// TIA Portal V19 export
// export: Created 2026-10-15T10:10:37.1458644Z, ExportSetting WithDefaults, DisplayName Totally Integrated Automation Portal, DisplayVersion V19, DisplayName TIA Portal Openness, DisplayVersion V19, DisplayName TIA Portal Version Control Interface, DisplayVersion V19, DisplayName STEP 7 Professional, DisplayVersion V19, DisplayName STEP 7 Safety, DisplayVersion V19, DisplayName WinCC Basic/Comfort/Advanced, DisplayVersion V19, DisplayName WinCC Unified, DisplayVersion V19
FUNCTION "ROLL_ReadInputs" : Void   // FC36, SCL
{ S7_Optimized_Access := 'TRUE' }
VERSION : 0.1
// stored: AutoNumber true, IsIECCheckEnabled false, SetENOAutomatically false, UDAEnableTagReadback false
   VAR_TEMP
      "b" : Int;
      bit : Int;
   END_VAR
BEGIN

   // Confirmed four-station profile: absent optional inputs are zero.
   FOR #b := 119 TO 125 DO
       FOR #bit := 0 TO 7 DO
           "ROLL_IO".Input[#b, #bit] := FALSE;
       END_FOR;
   END_FOR;
   IF "ROLL_IO".PhysicalIoConfigured AND NOT "ROLL_IO".Simulation THEN
       "ROLL_IO".Input[0, 0] := "Tag__639276557951123186";
       "ROLL_IO".Input[0, 1] := "Tag__639276557952818668";
       "ROLL_IO".Input[0, 2] := "Tag__639276557952918398";
       "ROLL_IO".Input[0, 3] := "Tag__639276557952998183";
       "ROLL_IO".Input[0, 4] := "Tag__639276557953077986";
       "ROLL_IO".Input[0, 5] := "Tag__639276557953157762";
       "ROLL_IO".Input[0, 6] := "Tag__639276557953227573";
       "ROLL_IO".Input[0, 7] := "Tag__639276557953307358";
       "ROLL_IO".Input[1, 0] := "Tag__639276557953367206";
       "ROLL_IO".Input[1, 1] := "Tag__639276557953447409";
       "ROLL_IO".Input[1, 2] := "Tag__639276557953526828";
       "ROLL_IO".Input[1, 3] := "Tag__639276557953606562";
       "ROLL_IO".Input[1, 4] := "Tag__639276557953686353";
       "ROLL_IO".Input[1, 5] := "Tag__639276557953766129";
       "ROLL_IO".Input[1, 6] := "Tag__639276557953835956";
       "ROLL_IO".Input[1, 7] := "Tag__639276557953915729";
       "ROLL_IO".Input[2, 0] := "Tag__639276557953985541";
       "ROLL_IO".Input[2, 1] := "Tag__639276557954055362";
       "ROLL_IO".Input[2, 2] := "Tag__639276557954135145";
       "ROLL_IO".Input[2, 3] := "Tag__639276557954204958";
       "ROLL_IO".Input[2, 4] := "Tag__639276557954284740";
       "ROLL_IO".Input[2, 5] := "Tag__639276557954354781";
       "ROLL_IO".Input[2, 6] := "Tag__639276557954434344";
       "ROLL_IO".Input[2, 7] := "Tag__639276557954494175";
       "ROLL_IO".Input[3, 0] := "Tag__639276557954554015";
       "ROLL_IO".Input[3, 1] := "Tag__639276557954604247";
       "ROLL_IO".Input[3, 2] := "Tag__639276557954663730";
       "ROLL_IO".Input[3, 3] := "Tag__639276557954723560";
       "ROLL_IO".Input[3, 4] := "Tag__639276557954773427";
       "ROLL_IO".Input[3, 5] := "Tag__639276557954833268";
       "ROLL_IO".Input[3, 6] := "Tag__639276557954893102";
       "ROLL_IO".Input[3, 7] := "Tag__639276557954953006";
       "ROLL_IO".Input[4, 0] := "Tag__639276557955012796";
       "ROLL_IO".Input[4, 1] := "Tag__639276557955062653";
       "ROLL_IO".Input[4, 2] := "Tag__639276557955122494";
       "ROLL_IO".Input[4, 3] := "Tag__639276557955182529";
       "ROLL_IO".Input[4, 4] := "Tag__639276557955242183";
       "ROLL_IO".Input[4, 5] := "Tag__639276557955302013";
       "ROLL_IO".Input[4, 6] := "Tag__639276557955362031";
       "ROLL_IO".Input[4, 7] := "Tag__639276557955411719";
       "ROLL_IO".Input[5, 0] := "Tag__639276557955481879";
       "ROLL_IO".Input[5, 1] := "Tag__639276557955541374";
       "ROLL_IO".Input[5, 2] := "Tag__639276557955601431";
       "ROLL_IO".Input[5, 3] := "Tag__639276557955661053";
       "ROLL_IO".Input[5, 4] := "Tag__639276557955710919";
       "ROLL_IO".Input[5, 5] := "Tag__639276557955770760";
       "ROLL_IO".Input[5, 6] := "Tag__639276557955820633";
       "ROLL_IO".Input[5, 7] := "Tag__639276557955880472";
       "ROLL_IO".Input[6, 0] := "Tag__639276557955940421";
       "ROLL_IO".Input[6, 1] := "Tag__639276557955990183";
       "ROLL_IO".Input[6, 2] := "Tag__639276557956050021";
       "ROLL_IO".Input[6, 3] := "Tag__639276557956099878";
       "ROLL_IO".Input[6, 4] := "Tag__639276557956149744";
       "ROLL_IO".Input[6, 5] := "Tag__639276557956209908";
       "ROLL_IO".Input[6, 6] := "Tag__639276557956259702";
       "ROLL_IO".Input[6, 7] := "Tag__639276557956319298";
       "ROLL_IO".Input[7, 0] := "Tag__639276557956369159";
       "ROLL_IO".Input[7, 1] := "Tag__639276557956419023";
       "ROLL_IO".Input[7, 2] := "Tag__639276557956479295";
       "ROLL_IO".Input[7, 3] := "Tag__639276557956528731";
       "ROLL_IO".Input[7, 4] := "Tag__639276557956578596";
       "ROLL_IO".Input[7, 5] := "Tag__639276557956638440";
       "ROLL_IO".Input[7, 6] := "Tag__639276557956698277";
       "ROLL_IO".Input[7, 7] := "Tag__639276557956758124";
       "ROLL_IO".Input[8, 0] := "Tag__639276557956808017";
       "ROLL_IO".Input[8, 1] := "Tag__639276557956867823";
       "ROLL_IO".Input[8, 2] := "Tag__639276557956917689";
       "ROLL_IO".Input[8, 3] := "Tag__639276557956977678";
       "ROLL_IO".Input[8, 4] := "Tag__639276557957037371";
       "ROLL_IO".Input[8, 5] := "Tag__639276557957087293";
       "ROLL_IO".Input[8, 6] := "Tag__639276557957147084";
       "ROLL_IO".Input[8, 7] := "Tag__639276557957196942";
       "ROLL_IO".Input[9, 0] := "Tag__639276557957256782";
       "ROLL_IO".Input[9, 1] := "Tag__639276557957316622";
       "ROLL_IO".Input[9, 2] := "Tag__639276557957366490";
       "ROLL_IO".Input[9, 3] := "Tag__639276557957426337";
       "ROLL_IO".Input[9, 4] := "Tag__639276557957476206";
       "ROLL_IO".Input[9, 5] := "Tag__639276557957526061";
       "ROLL_IO".Input[9, 6] := "Tag__639276557957586243";
       "ROLL_IO".Input[9, 7] := "Tag__639276557957645746";
       "ROLL_IO".Input[10, 0] := "Tag__639276557957705582";
       "ROLL_IO".Input[10, 1] := "Tag__639276557957755449";
       "ROLL_IO".Input[10, 2] := "Tag__639276557957805314";
       "ROLL_IO".Input[10, 3] := "Tag__639276557957865154";
       "ROLL_IO".Input[10, 4] := "Tag__639276557957915021";
       "ROLL_IO".Input[10, 5] := "Tag__639276557957964888";
       "ROLL_IO".Input[10, 6] := "Tag__639276557958024728";
       "ROLL_IO".Input[10, 7] := "Tag__639276557958074957";
       "ROLL_IO".Input[11, 0] := "Tag__639276557958124460";
       "ROLL_IO".Input[11, 1] := "Tag__639276557958184301";
       "ROLL_IO".Input[11, 2] := "Tag__639276557958234167";
       "ROLL_IO".Input[11, 3] := "Tag__639276557958294016";
       "ROLL_IO".Input[11, 4] := "Tag__639276557958343874";
       "ROLL_IO".Input[11, 5] := "Tag__639276557958393749";
       "ROLL_IO".Input[11, 6] := "Tag__639276557958453636";
       "ROLL_IO".Input[11, 7] := "Tag__639276557958503448";
       "ROLL_IO".Input[12, 0] := "Tag__639276557958553313";
       "ROLL_IO".Input[12, 1] := "Tag__639276557958613155";
       "ROLL_IO".Input[12, 2] := "Tag__639276557958663020";
       "ROLL_IO".Input[12, 3] := "Tag__639276557958712886";
       "ROLL_IO".Input[12, 4] := "Tag__639276557958772727";
       "ROLL_IO".Input[12, 5] := "Tag__639276557958822593";
       "ROLL_IO".Input[12, 6] := "Tag__639276557958902547";
       "ROLL_IO".Input[12, 7] := "Tag__639276557958962223";
       "ROLL_IO".Input[13, 0] := "Tag__639276557959022060";
       "ROLL_IO".Input[13, 1] := "Tag__639276557959071925";
       "ROLL_IO".Input[13, 2] := "Tag__639276557959131766";
       "ROLL_IO".Input[13, 3] := "Tag__639276557959191606";
       "ROLL_IO".Input[13, 4] := "Tag__639276557959251774";
       "ROLL_IO".Input[13, 5] := "Tag__639276557959311297";
       "ROLL_IO".Input[13, 6] := "Tag__639276557959371125";
       "ROLL_IO".Input[13, 7] := "Tag__639276557959430966";
       "ROLL_IO".Input[14, 0] := "Tag__639276557959490814";
       "ROLL_IO".Input[14, 1] := "Tag__639276557959540672";
       "ROLL_IO".Input[14, 2] := "Tag__639276557959600839";
       "ROLL_IO".Input[14, 3] := "Tag__639276557959650385";
       "ROLL_IO".Input[14, 4] := "Tag__639276557959710219";
       "ROLL_IO".Input[14, 5] := "Tag__639276557959760095";
       "ROLL_IO".Input[14, 6] := "Tag__639276557959809951";
       "ROLL_IO".Input[14, 7] := "Tag__639276557959869792";
       "ROLL_IO".Input[15, 0] := "Tag__639276557959929638";
       "ROLL_IO".Input[15, 1] := "Tag__639276557959979499";
       "ROLL_IO".Input[15, 2] := "Tag__639276557960039343";
       "ROLL_IO".Input[15, 3] := "Tag__639276557960089204";
       "ROLL_IO".Input[15, 4] := "Tag__639276557960139071";
       "ROLL_IO".Input[15, 5] := "Tag__639276557960198912";
       "ROLL_IO".Input[15, 6] := "Tag__639276557960248790";
       "ROLL_IO".Input[15, 7] := "Tag__639276557960308618";
   END_IF;
END_FUNCTION
